Fanuc KAREL source: kf00040.KL

-- PROVISIONAL review KL for V1013-1; original PC SHA256 099cf652ca62e00fa99c3c0c8d792c8bd41419715c847103dbb13016cd6fd3f6
-- Incomplete behavior may be omitted. Consult companion uncertainty JSON. Do not deploy.
PROGRAM KF00040
%NOLOCKGROUP
VAR
  I : INTEGER
  J : INTEGER
  X : REAL
  Y : REAL
  B : BOOLEAN
  C : BOOLEAN
  TXT : STRING[80]
  TXT2 : STRING[80]
  STATUS : INTEGER
-- UNRESOLVED_DECL AI type=002010
-- UNRESOLVED_DECL BI type=002010
-- UNRESOLVED_DECL P type=000102
-- UNRESOLVED_DECL JP type=000199
-- UNRESOLVED_DECL PF type=000101
-- UNRESOLVED_DECL V1 type=000013
-- UNRESOLVED_DECL V2 type=000013
BEGIN
  -- UNRESOLVED_PC offsets 5-19; opcodes 3F,75
  -- UNRESOLVED_PC offsets 24-36; opcodes 73,75
  -- UNRESOLVED_PC offsets 41-45; opcodes 7F
END KF00040
